TYPE ST_MixProof_state :
STRUCT
	sName: STRING;
	bUpper: BOOL;
	bLower: BOOL;
	bRunning: BOOL;
	bDone: BOOL;

END_STRUCT
END_TYPE

(* stored: Version 1.1.0.1, ProductVersion 3.1.4024.13
   DUT ST_MixProof_state: Id {a1caa6fd-e6aa-4e55-ab79-2047e0dc9fac} *)
